Fanuc KAREL source: KT00199.KL

PROGRAM KT00199
%NOLOCKGROUP
VAR
  B1: BOOLEAN
  H2: ARRAY[2] OF SHORT
  OUT: BOOLEAN
BEGIN
  B1 = TRUE
    H2[1] = 3
  OUT = B1 AND H2[1]
END KT00199
